(* IEC 61131-3 sources: rusty/compiler/plc_cfc/fixtures/execution_control/valid/enable_from_block, 2 files *)

(* ---- counter.st ---- *)
FUNCTION_BLOCK counter
VAR_INPUT
    in : DINT;
END_VAR
VAR_OUTPUT
    out : DINT;
END_VAR
    out := out + in;
END_FUNCTION_BLOCK

(* ---- gate.st ---- *)
FUNCTION_BLOCK gate
VAR_OUTPUT
    ok : BOOL;
END_VAR
    ok := TRUE;
END_FUNCTION_BLOCK
